PROGRAM main
VAR
	M_EStop_Latch : bool;
	M_GarageFull : bool;
	M_Crossing_Occ : bool;
	Failsafe_Cond : bool;
	Failsafe_Prev : bool;
	Failsafe_Trip : bool;
	EndL_Stable : bool;
	EndR_Stable : bool;
	Xing_Latched : bool;
	Xing_EnteredA : bool;
	Xing_EnteredB : bool;
	GarageL_Deb : TON;
	GarageR_Deb : TON;
	Xing_Clear_Delay : TOF;
	TRIP_CM : int := 5;
	Power_FB AT %IX100.0 : bool;
	EStop_Button AT %IX100.1 : bool;
	VR_OK AT %IX100.2 : bool;
	IR_CrossA AT %IX100.3 : bool;
	IR_CrossB AT %IX100.4 : bool;
	IR_EndL AT %IX100.5 : bool;
	IR_EndR AT %IX100.6 : bool;
	Ultrasonic_Dist AT %IW103 : int;
	Track_Power_Cmd AT %QX100.0 : bool;
	Buzzer_Cmd AT %QX100.1 : bool;
	J1_Angle AT %QW100 : int;
	J2_Angle AT %QW101 : int;
	Crossing_Gate AT %QW102 : int;
	LED_Mode AT %QW103 : int;
	Failsafe_Servo AT %QW104 : int;
	LCD1_Code AT %QW105 : int;
	LCD2_Code AT %QW106 : int;
	LCD3_Code AT %QW107 : int;
	Reset_Cmd AT %QX80.0 : bool;
	Run_Cmd AT %QX80.1 : bool;
	EStop_SW AT %QX80.2 : bool;
	Manual_Mode AT %QX80.3 : bool;
	J1_Cmd AT %QX80.4 : bool;
	J2_Cmd AT %QX80.5 : bool;
END_VAR

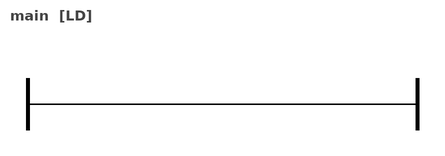
(* LD diagram, written out as Structured Text *)
END_PROGRAM
